(* IEC 61131-3 sources: s7-to-codesys/tests/POUs/S7Compat/FB_S7Tp_Test, 4 files *)

(* ---- FB_S7Tp_Test.decl.st ---- *)
// Назначение: набор тестов CfUnit (coUnit 1.2.0.0) для FB_S7Tp слоя совместимости S7Compat:
//             импульс по фронту IN длительностью PT, порог PT, ET после импульса и при IN = FALSE,
//             фронты во время импульса, совпадение со Standard.TP в реальном времени.
//             Ожидаемые значения — по семантике МЭК 61131-3 и S7 (описание в объявлении блока), а
//             не по результату реализации. Моделируемое время — GVL_S7Clock (тест включает и
//             выключает его сам). Экземпляр набора объявляется в PRG_Tests.
// Автор:      kr0nsch
// Версия:     0.1.0
// Документ:   docs/methodology.md, раздел «Проверка поведения: время в тестах»
FUNCTION_BLOCK FB_S7Tp_Test EXTENDS coUnit.FB_TestSuite
VAR
    // MatchesStandardInRealTime: состояние между циклами (тест идёт несколько циклов)
    fbRtCompat : FB_S7Tp;              // проверяемый таймер S7Compat
    fbRtStandard : TP;               // эталон — таймер CODESYS Standard
    xRtStarted : BOOL;              // момент начала зафиксирован
    xRtDone : BOOL;                 // тест завершён
    xRtIn : BOOL;                   // общий вход IN
    xRtSawQ : BOOL;                 // Standard Q хотя бы раз был TRUE
    tRtStart : TIME;                // время начала теста (F_S7Now() = TIME())
    tRtElapsed : TIME;              // прошло с начала теста
    tRtEtDiff : TIME;               // |ET S7Compat - ET Standard|
    tRtEtToPt : TIME;               // PT - ET Standard (близость к порогу)
    iRtMismatches : INT;            // циклов с расхождением
END_VAR
VAR CONSTANT
    T_RT_PT : TIME := T#200MS;      // PT обоих таймеров
    T_RT_DURATION : TIME := T#700MS;  // длительность теста
    T_RT_TOL : TIME := T#5MS;       // допуск ET: таймеры читают TIME() в разные моменты цикла
END_VAR

(* ---- MatchesStandardInRealTime.method.impl.st ---- *)
coUnit.TEST('MatchesStandardInRealTime');
IF NOT xRtDone THEN
    IF NOT xRtStarted THEN
        xRtStarted := TRUE;
        tRtStart := F_S7Now();  // xSimulation = FALSE: время ПЛК, как TIME()
    END_IF
    tRtElapsed := F_S7Now() - tRtStart;
    xRtIn := (tRtElapsed < T#100MS) OR (tRtElapsed >= T#150MS AND tRtElapsed < T#500MS);
    fbRtCompat(IN := xRtIn, PT := T_RT_PT);
    fbRtStandard(IN := xRtIn, PT := T_RT_PT);
    IF fbRtCompat.ET >= fbRtStandard.ET THEN
        tRtEtDiff := fbRtCompat.ET - fbRtStandard.ET;
    ELSE
        tRtEtDiff := fbRtStandard.ET - fbRtCompat.ET;
    END_IF
    tRtEtToPt := T_RT_PT - fbRtStandard.ET;  // ET <= PT
    IF tRtEtDiff > T_RT_TOL OR (fbRtCompat.Q <> fbRtStandard.Q AND tRtEtToPt > T_RT_TOL) THEN
        iRtMismatches := iRtMismatches + 1;
    END_IF
    xRtSawQ := xRtSawQ OR fbRtStandard.Q;
    IF tRtElapsed >= T_RT_DURATION THEN
        xRtDone := TRUE;
        AssertEquals_INT(Expected := 0, Actual := iRtMismatches, Message := 'FB_S7Tp vs TP: mismatching cycles');
        AssertTrue(Condition := xRtSawQ, Message := 'FB_S7Tp vs TP: Standard Q never TRUE, test did not run');
    END_IF
END_IF
IF xRtDone THEN
    coUnit.TEST_FINISHED();
END_IF

(* ---- PulseOnRisingEdge.method.decl.st ---- *)
// фронт IN на 0 мс, PT = 1 с: Q = TRUE до 999 мс, FALSE на 1000 мс; ET = PT, пока IN = TRUE; 0 при IN = FALSE.
METHOD PRIVATE PulseOnRisingEdge
VAR
    fbDut : FB_S7Tp;       // проверяемый таймер (новый экземпляр на каждый вызов метода)
END_VAR

(* ---- RetriggerIgnored.method.decl.st ---- *)
// фронт IN во время импульса не продлевает его; спад IN во время импульса его не обрывает.
METHOD PRIVATE RetriggerIgnored
VAR
    fbDut : FB_S7Tp;       // проверяемый таймер (новый экземпляр на каждый вызов метода)
END_VAR
